// Mitsubishi GX Works2 project: AGV_IOCHECK   PLC: Q03UD

PROGRAM IOCHECK
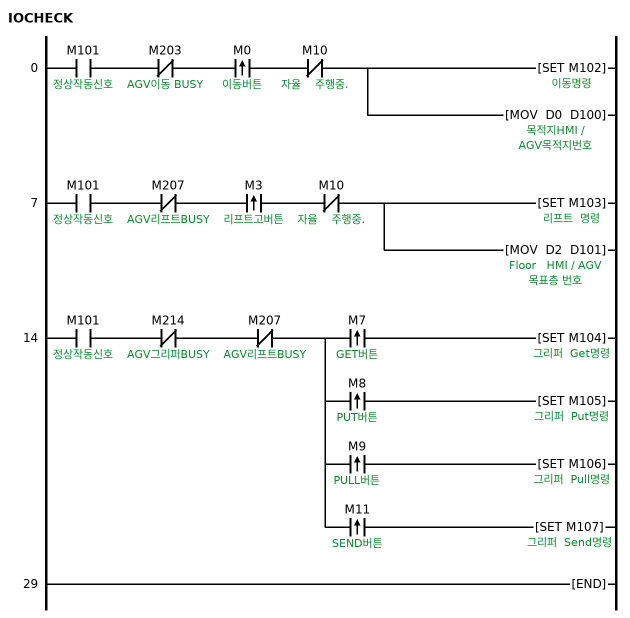
0     LD      M101  ; 정상작동신호
      ANI     M203  ; AGV이동 BUSY
      ANDP    M0  ; 이동버튼
      ANI     M10  ; 자율    주행중.
      SET     M102  ; 이동명령
      MOV     D0 D100  ; 목적지HMI / AGV목적지번호
7     LD      M101  ; 정상작동신호
      ANI     M207  ; AGV리프트BUSY
      ANDP    M3  ; 리프트고버튼
      ANI     M10  ; 자율    주행중.
      SET     M103  ; 리프트  명령
      MOV     D2 D101  ; Floor   HMI / AGV 목표층 번호
14    LD      M101  ; 정상작동신호
      ANI     M214  ; AGV그리퍼BUSY
      ANI     M207  ; AGV리프트BUSY
      MPS
      ANDP    M7  ; GET버튼
      SET     M104  ; 그리퍼  Get명령
      MRD
      ANDP    M8  ; PUT버튼
      SET     M105  ; 그리퍼  Put명령
      MRD
      ANDP    M9  ; PULL버튼
      SET     M106  ; 그리퍼  Pull명령
      MPP
      ANDP    M11  ; SEND버튼
      SET     M107  ; 그리퍼  Send명령
29    END
END_PROGRAM

PROGRAM MAIN
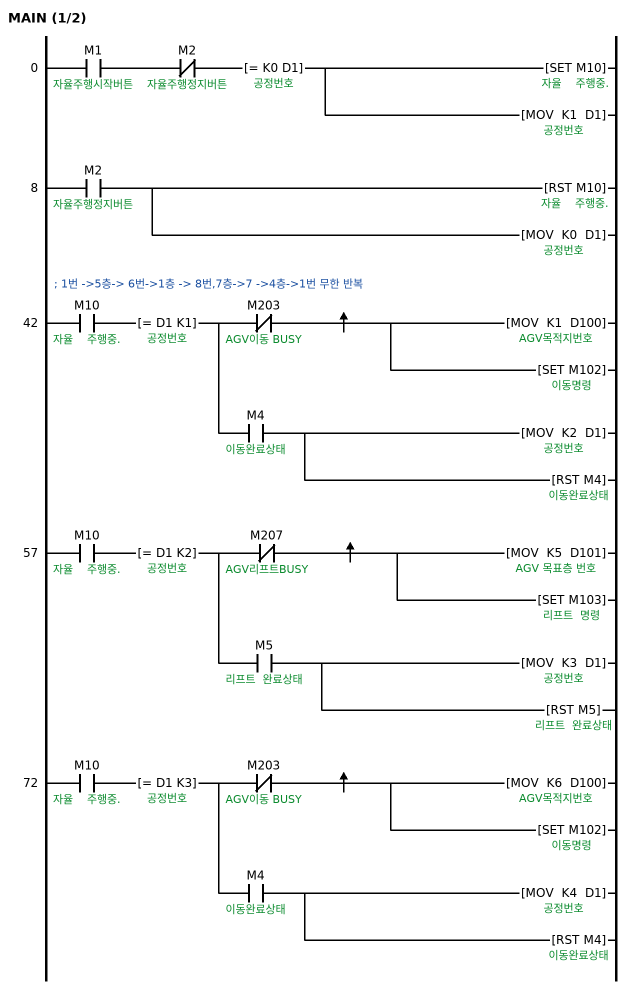
0     LD      M1  ; 자율주행시작버튼
      ANI     M2  ; 자율주행정지버튼
      AND=    K0 D1  ; 공정번호
      SET     M10  ; 자율    주행중.
      MOV     K1 D1
8     LD      M2  ; 자율주행정지버튼
      RST     M10  ; 자율    주행중.
      MOV     K0 D1
; 1번 ->5층-> 6번->1층 -> 8번,7층->7 ->4층->1번 무한 반복
42    LD      M10  ; 자율    주행중.
      AND=    D1 K1  ; 공정번호
      MPS
      ANI     M203  ; AGV이동 BUSY
      MEP
      MOV     K1 D100  ; AGV목적지번호
      SET     M102  ; 이동명령
      MPP
      AND     M4  ; 이동완료상태
      MOV     K2 D1
      RST     M4  ; 이동완료상태
57    LD      M10  ; 자율    주행중.
      AND=    D1 K2  ; 공정번호
      MPS
      ANI     M207  ; AGV리프트BUSY
      MEP
      MOV     K5 D101  ; AGV 목표층 번호
      SET     M103  ; 리프트  명령
      MPP
      AND     M5  ; 리프트  완료상태
      MOV     K3 D1
      RST     M5  ; 리프트  완료상태
72    LD      M10  ; 자율    주행중.
      AND=    D1 K3  ; 공정번호
      MPS
      ANI     M203  ; AGV이동 BUSY
      MEP
      MOV     K6 D100
      SET     M102  ; 이동명령
      MPP
      AND     M4  ; 이동완료상태
      MOV     K4 D1
      RST     M4  ; 이동완료상태
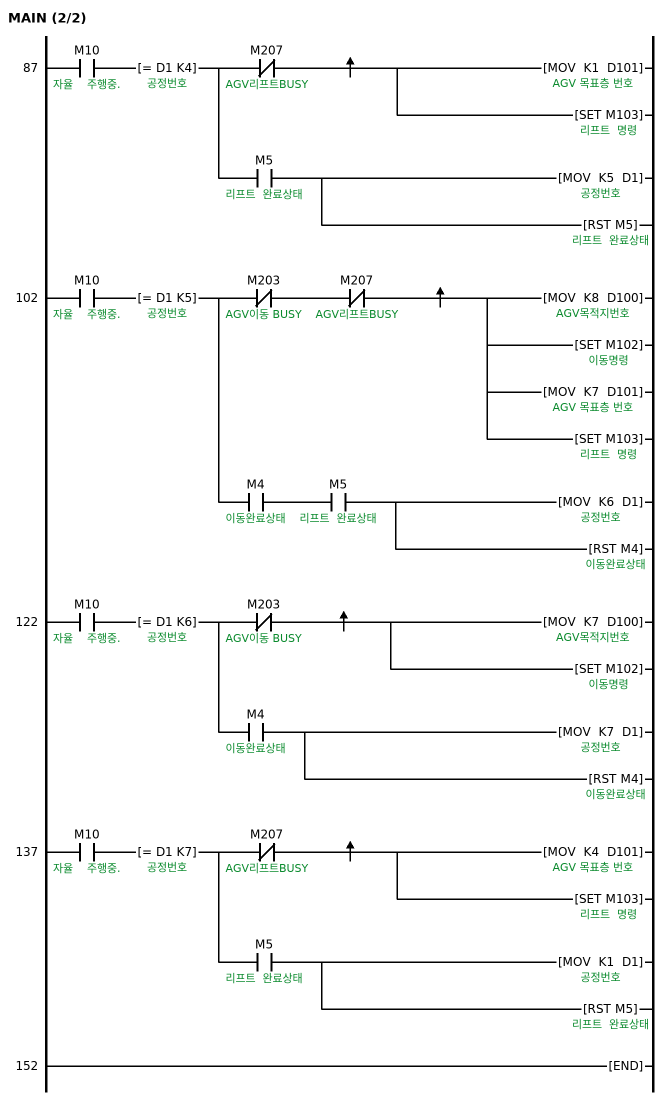
87    LD      M10  ; 자율    주행중.
      AND=    D1 K4  ; 공정번호
      MPS
      ANI     M207  ; AGV리프트BUSY
      MEP
      MOV     K1 D101
      SET     M103  ; 리프트  명령
      MPP
      AND     M5  ; 리프트  완료상태
      MOV     K5 D1
      RST     M5  ; 리프트  완료상태
102   LD      M10  ; 자율    주행중.
      AND=    D1 K5  ; 공정번호
      MPS
      ANI     M203  ; AGV이동 BUSY
      ANI     M207  ; AGV리프트BUSY
      MEP
      MOV     K8 D100
      SET     M102  ; 이동명령
      MOV     K7 D101
      SET     M103  ; 리프트  명령
      MPP
      AND     M4  ; 이동완료상태
      AND     M5  ; 리프트  완료상태
      MOV     K6 D1
      RST     M4  ; 이동완료상태
122   LD      M10  ; 자율    주행중.
      AND=    D1 K6  ; 공정번호
      MPS
      ANI     M203  ; AGV이동 BUSY
      MEP
      MOV     K7 D100
      SET     M102  ; 이동명령
      MPP
      AND     M4  ; 이동완료상태
      MOV     K7 D1
      RST     M4  ; 이동완료상태
137   LD      M10  ; 자율    주행중.
      AND=    D1 K7  ; 공정번호
      MPS
      ANI     M207  ; AGV리프트BUSY
      MEP
      MOV     K4 D101
      SET     M103  ; 리프트  명령
      MPP
      AND     M5  ; 리프트  완료상태
      MOV     K1 D1
      RST     M5  ; 리프트  완료상태
152   END
END_PROGRAM

PROGRAM INPUT
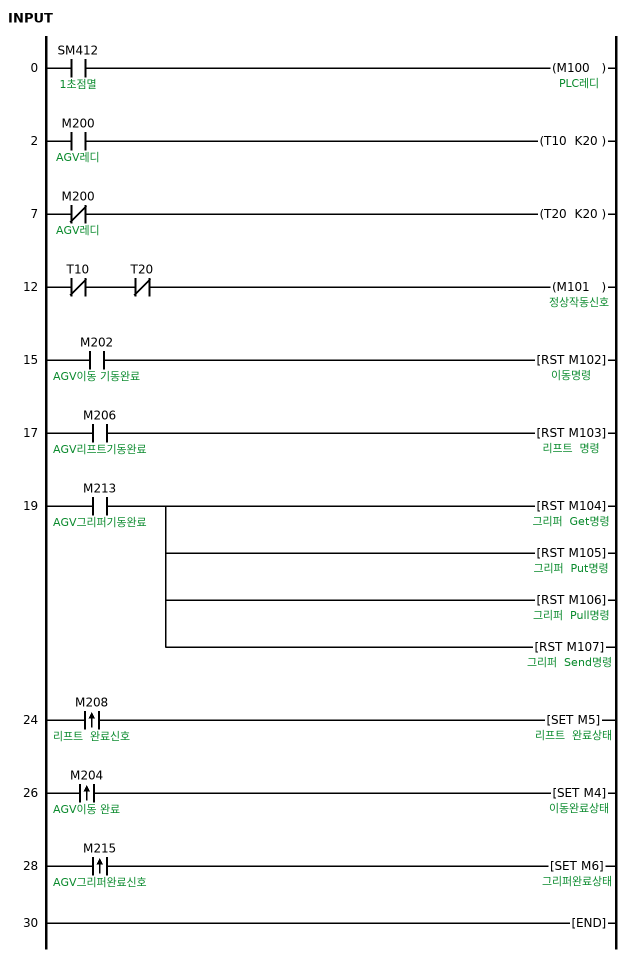
0     LD      SM412  ; 1초점멸
      OUT     M100  ; PLC레디
2     LD      M200  ; AGV레디
      OUT     T10 K20
7     LDI     M200  ; AGV레디
      OUT     T20 K20
12    LDI     T10
      ANI     T20
      OUT     M101  ; 정상작동신호
15    LD      M202  ; AGV이동 기동완료
      RST     M102  ; 이동명령
17    LD      M206  ; AGV리프트기동완료
      RST     M103  ; 리프트  명령
19    LD      M213  ; AGV그리퍼기동완료
      RST     M104  ; 그리퍼  Get명령
      RST     M105  ; 그리퍼  Put명령
      RST     M106  ; 그리퍼  Pull명령
      RST     M107  ; 그리퍼  Send명령
24    LDP     M208  ; 리프트  완료신호
      SET     M5  ; 리프트  완료상태
26    LDP     M204  ; AGV이동 완료
      SET     M4  ; 이동완료상태
28    LDP     M215  ; AGV그리퍼완료신호
      SET     M6  ; 그리퍼완료상태
30    END
END_PROGRAM

PROGRAM OUTPUT
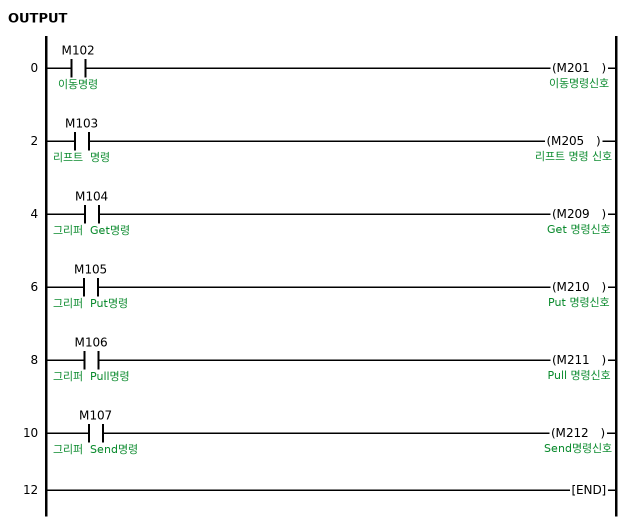
0     LD      M102  ; 이동명령
      OUT     M201  ; 이동명령신호
2     LD      M103  ; 리프트  명령
      OUT     M205  ; 리프트 명령 신호
4     LD      M104  ; 그리퍼  Get명령
      OUT     M209  ; Get 명령신호
6     LD      M105  ; 그리퍼  Put명령
      OUT     M210  ; Put 명령신호
8     LD      M106  ; 그리퍼  Pull명령
      OUT     M211  ; Pull 명령신호
10    LD      M107  ; 그리퍼  Send명령
      OUT     M212  ; Send명령신호
12    END
END_PROGRAM

PROGRAM MAIN2
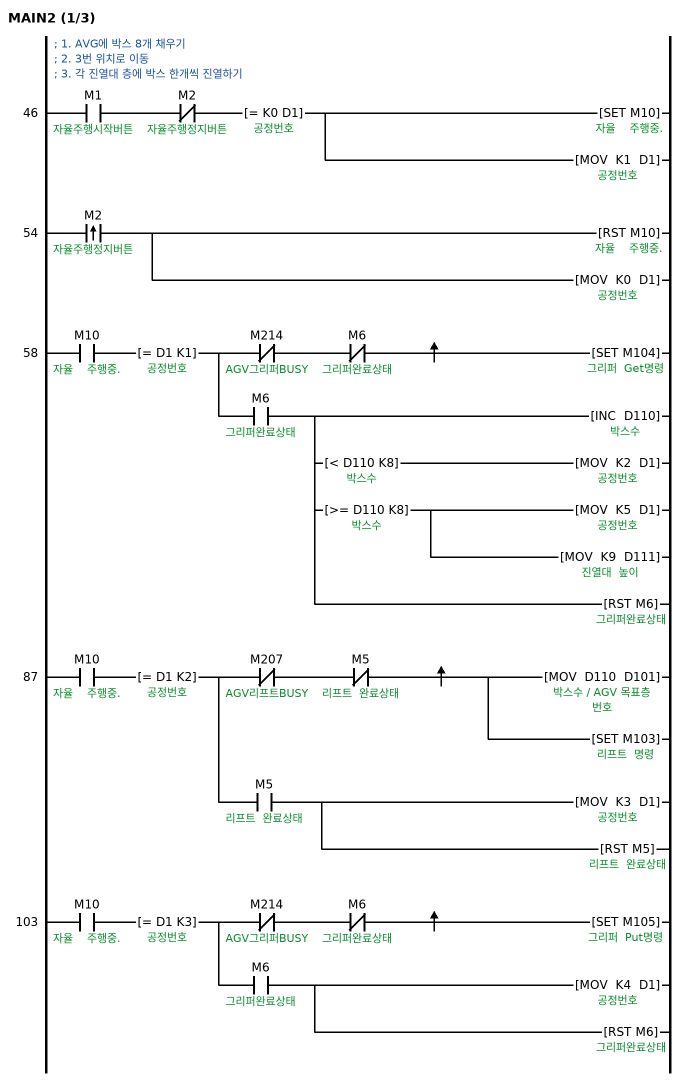
; 1. AVG에 박스 8개 채우기
; 2. 3번 위치로 이동
; 3. 각 진열대 층에 박스 한개씩 진열하기
46    LD      M1  ; 자율주행시작버튼
      ANI     M2  ; 자율주행정지버튼
      AND=    K0 D1  ; 공정번호
      SET     M10  ; 자율    주행중.
      MOV     K1 D1
54    LDP     M2  ; 자율주행정지버튼
      RST     M10  ; 자율    주행중.
      MOV     K0 D1
58    LD      M10  ; 자율    주행중.
      AND=    D1 K1  ; 공정번호
      MPS
      ANI     M214  ; AGV그리퍼BUSY
      ANI     M6  ; 그리퍼완료상태
      MEP
      SET     M104  ; 그리퍼  Get명령
      MPP
      AND     M6  ; 그리퍼완료상태
      INC     D110  ; 박스수
      MPS
      AND<    D110 K8  ; 박스수
      MOV     K2 D1
      MRD
      AND>=   D110 K8  ; 박스수
      MOV     K5 D1
      MOV     K9 D111  ; 진열대  높이
      MPP
      RST     M6  ; 그리퍼완료상태
87    LD      M10  ; 자율    주행중.
      AND=    D1 K2  ; 공정번호
      MPS
      ANI     M207  ; AGV리프트BUSY
      ANI     M5  ; 리프트  완료상태
      MEP
      MOV     D110 D101  ; AGV 목표층 번호
      SET     M103  ; 리프트  명령
      MPP
      AND     M5  ; 리프트  완료상태
      MOV     K3 D1
      RST     M5  ; 리프트  완료상태
103   LD      M10  ; 자율    주행중.
      AND=    D1 K3  ; 공정번호
      MPS
      ANI     M214  ; AGV그리퍼BUSY
      ANI     M6  ; 그리퍼완료상태
      MEP
      SET     M105  ; 그리퍼  Put명령
      MPP
      AND     M6  ; 그리퍼완료상태
      MOV     K4 D1
      RST     M6  ; 그리퍼완료상태
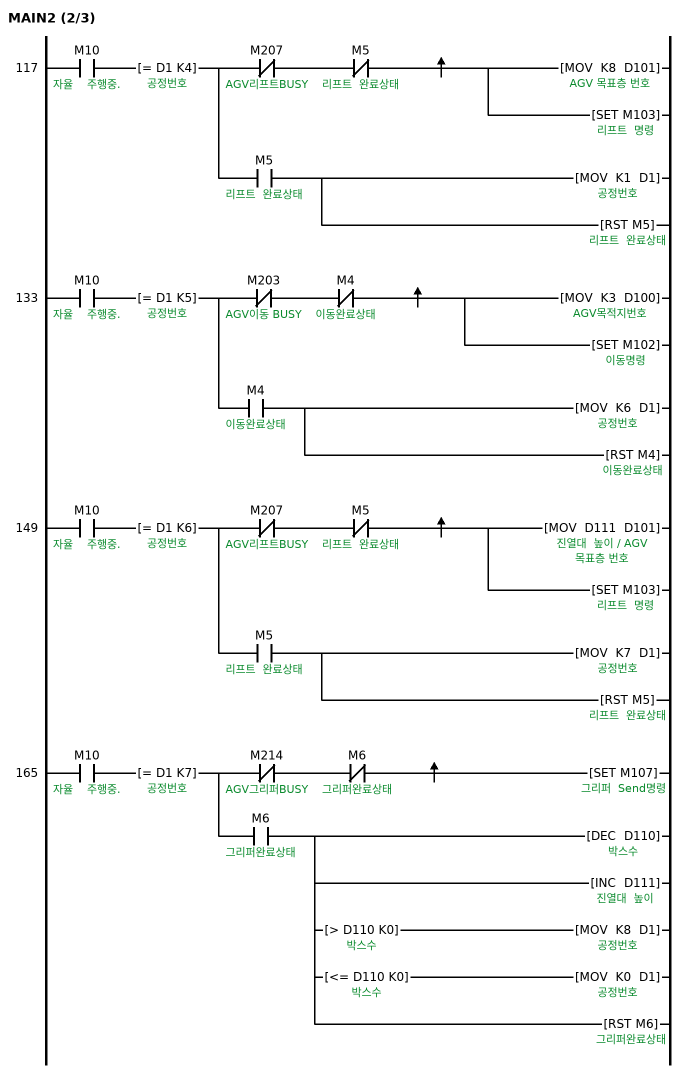
117   LD      M10  ; 자율    주행중.
      AND=    D1 K4  ; 공정번호
      MPS
      ANI     M207  ; AGV리프트BUSY
      ANI     M5  ; 리프트  완료상태
      MEP
      MOV     K8 D101
      SET     M103  ; 리프트  명령
      MPP
      AND     M5  ; 리프트  완료상태
      MOV     K1 D1
      RST     M5  ; 리프트  완료상태
133   LD      M10  ; 자율    주행중.
      AND=    D1 K5  ; 공정번호
      MPS
      ANI     M203  ; AGV이동 BUSY
      ANI     M4  ; 이동완료상태
      MEP
      MOV     K3 D100  ; AGV목적지번호
      SET     M102  ; 이동명령
      MPP
      AND     M4  ; 이동완료상태
      MOV     K6 D1
      RST     M4  ; 이동완료상태
149   LD      M10  ; 자율    주행중.
      AND=    D1 K6  ; 공정번호
      MPS
      ANI     M207  ; AGV리프트BUSY
      ANI     M5  ; 리프트  완료상태
      MEP
      MOV     D111 D101
      SET     M103  ; 리프트  명령
      MPP
      AND     M5  ; 리프트  완료상태
      MOV     K7 D1
      RST     M5  ; 리프트  완료상태
165   LD      M10  ; 자율    주행중.
      AND=    D1 K7  ; 공정번호
      MPS
      ANI     M214  ; AGV그리퍼BUSY
      ANI     M6  ; 그리퍼완료상태
      MEP
      SET     M107  ; 그리퍼  Send명령
      MPP
      AND     M6  ; 그리퍼완료상태
      DEC     D110
      INC     D111
      MPS
      AND>    D110 K0  ; 박스수
      MOV     K8 D1
      MRD
      AND<=   D110 K0  ; 박스수
      MOV     K0 D1
      MPP
      RST     M6  ; 그리퍼완료상태
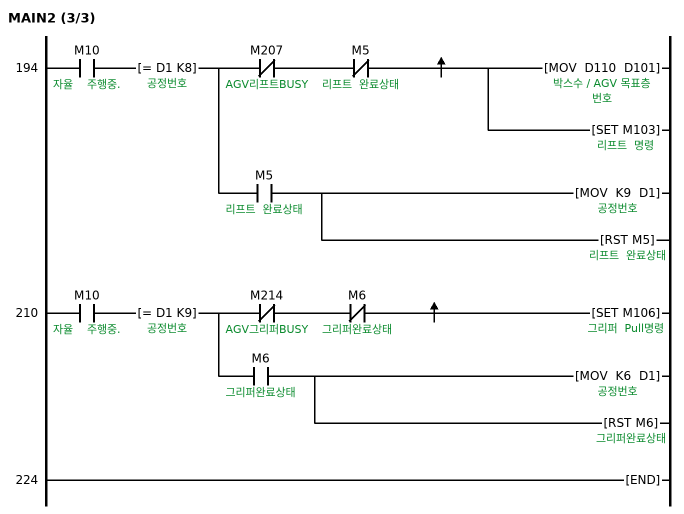
194   LD      M10  ; 자율    주행중.
      AND=    D1 K8  ; 공정번호
      MPS
      ANI     M207  ; AGV리프트BUSY
      ANI     M5  ; 리프트  완료상태
      MEP
      MOV     D110 D101
      SET     M103  ; 리프트  명령
      MPP
      AND     M5  ; 리프트  완료상태
      MOV     K9 D1
      RST     M5  ; 리프트  완료상태
210   LD      M10  ; 자율    주행중.
      AND=    D1 K9  ; 공정번호
      MPS
      ANI     M214  ; AGV그리퍼BUSY
      ANI     M6  ; 그리퍼완료상태
      MEP
      SET     M106  ; 그리퍼  Pull명령
      MPP
      AND     M6  ; 그리퍼완료상태
      MOV     K6 D1
      RST     M6  ; 그리퍼완료상태
224   END
END_PROGRAM

// device comments not shown above
M17  ; 그리퍼  Send명령
